(* IEC 61131-3 sources: plcassist-cli/packages/volt-lsp-iec/test-corpus/lenze-mid/Device/Plc Logic/Application/A71_LocalSources/CamControls/Pulse, 2 files *)

(* ---- fc_CamC_CP_Base.fun ---- *)
FUNCTION fc_CamC_CP_Base : BOOL
VAR_INPUT
	iEN					: BOOL;
	iStartCam			: INT;
	iMachinePosition 	: INT;
	iResetFlag			: BOOL;
END_VAR
VAR_OUTPUT

END_VAR
VAR
	tBool: BOOL;

END_VAR
VAR_IN_OUT
	ioAuxOneShot: BOOL;
END_VAR

NETWORK 0 LD
  LET en1 := ;
  IF en1 THEN (iMachinePosition >= iStartCam); END_IF
  tBool := (en1 AND NOT iResetFlag AND iEN);
END_NETWORK
NETWORK 1 LD
  fc_CamC_CP_Base := (tbool AND NOT ioAuxOneShot);
END_NETWORK
NETWORK 2 LD
  ioAuxOneShot := tbool;
END_NETWORK

END_FUNCTION

(* ---- fc_CamC_CP_UDT.fun ---- *)
FUNCTION fc_CamC_CP_UDT : BOOL
VAR_INPUT
	iEN						: BOOL;
	iMachinePosition		: INT;
	iResetFlag				: BOOL;

END_VAR
VAR_OUTPUT

END_VAR
VAR

END_VAR
VAR_IN_OUT
	ioPulse	: UDT_CamPulse;
END_VAR

NETWORK 0 LD
  LET en1 := ;
  IF en1 THEN ioPulse.MachinePos_HMI := MOVE(iMachinePosition); END_IF
END_NETWORK
NETWORK 1 LD
  LET g1 := fc_CamC_CP_Base(iEN, ioPulse.Start, iMachinePosition, iResetFlag, ioPulse.OSP);
  fc_CamC_CP_UDT := g1;
  ioPulse.Active := g1;
END_NETWORK

END_FUNCTION
